TYPE "ST_PressDemoReleaseConditions"
VERSION : 0.1
   STRUCT
      "ModeStartAirPressureOk" : Bool;
      "RamGuardClosed" : Bool;
      "RamSlideInside" : Bool;
      "RamDevicesHealthy" : Bool;
      "RamAirPressureOk" : Bool;
      "RamTwoHandHeld" : Bool;
   END_STRUCT;
END_TYPE
